// TIA Portal V19 export
// export: Created 2026-10-15T09:44:25.353626Z, ExportSetting WithDefaults, DisplayName Totally Integrated Automation Portal, DisplayVersion V19, DisplayName TIA Portal Openness, DisplayVersion V19, DisplayName TIA Portal Version Control Interface, DisplayVersion V19, DisplayName STEP 7 Professional, DisplayVersion V19, DisplayName STEP 7 Safety, DisplayVersion V19, DisplayName WinCC Basic/Comfort/Advanced, DisplayVersion V19, DisplayName WinCC Unified, DisplayVersion V19
FUNCTION "ROLL_WriteOutputs" : Void   // FC37, SCL
{ S7_Optimized_Access := 'TRUE' }
VERSION : 0.1
// stored: AutoNumber true, IsIECCheckEnabled false, SetENOAutomatically false, UDAEnableTagReadback false
   VAR_TEMP
      enabled : Bool;
   END_VAR
BEGIN

   IF "ROLL_IO".PhysicalIoConfigured THEN
       #enabled := "ROLL_IO".PhysicalOutputsEnabled AND NOT "ROLL_IO".Simulation AND NOT "ROLL_IO".ConversionFault;
       "Tag__639276542187652659" := #enabled AND "ROLL_IO".Output[16, 0];
       "Tag__639276542187732448" := #enabled AND "ROLL_IO".Output[16, 1];
       "Tag__639276542187792292" := #enabled AND "ROLL_IO".Output[16, 2];
       "Tag__639276542187852130" := #enabled AND "ROLL_IO".Output[16, 3];
       "Tag__639276542187911981" := #enabled AND "ROLL_IO".Output[16, 4];
       "Tag__639276542187972161" := #enabled AND "ROLL_IO".Output[16, 5];
       "Tag__639276542188021847" := #enabled AND "ROLL_IO".Output[16, 6];
       "Tag__639276542188081517" := #enabled AND "ROLL_IO".Output[16, 7];
       "Tag__639276542188141359" := #enabled AND "ROLL_IO".Output[17, 0];
       "Tag__639276542188191229" := #enabled AND "ROLL_IO".Output[17, 1];
       "Tag__639276542188251067" := #enabled AND "ROLL_IO".Output[17, 2];
       "Tag__639276542188320878" := #enabled AND "ROLL_IO".Output[17, 3];
       "Tag__639276542188410640" := #enabled AND "ROLL_IO".Output[17, 4];
       "Tag__639276542188520372" := #enabled AND "ROLL_IO".Output[17, 5];
       "Tag__639276542188610120" := #enabled AND "ROLL_IO".Output[17, 6];
       "Tag__639276542188699865" := #enabled AND "ROLL_IO".Output[17, 7];
       "Tag__639276542188769683" := #enabled AND "ROLL_IO".Output[18, 0];
       "Tag__639276542188839495" := #enabled AND "ROLL_IO".Output[18, 1];
       "Tag__639276542188899332" := #enabled AND "ROLL_IO".Output[18, 2];
       "Tag__639276542188969166" := #enabled AND "ROLL_IO".Output[18, 3];
       "Tag__639276542189049062" := #enabled AND "ROLL_IO".Output[18, 4];
       "Tag__639276542189108777" := #enabled AND "ROLL_IO".Output[18, 5];
       "Tag__639276542189178592" := #enabled AND "ROLL_IO".Output[18, 6];
       "Tag__639276542189258389" := #enabled AND "ROLL_IO".Output[18, 7];
       "Tag__639276542189338210" := #enabled AND "ROLL_IO".Output[19, 0];
       "Tag__639276542189407977" := #enabled AND "ROLL_IO".Output[19, 1];
       "Tag__639276542189488068" := #enabled AND "ROLL_IO".Output[19, 2];
       "Tag__639276542189557576" := #enabled AND "ROLL_IO".Output[19, 3];
       "Tag__639276542189627382" := #enabled AND "ROLL_IO".Output[19, 4];
       "Tag__639276542189697203" := #enabled AND "ROLL_IO".Output[19, 5];
       "Tag__639276542189767112" := #enabled AND "ROLL_IO".Output[19, 6];
       "Tag__639276542189836826" := #enabled AND "ROLL_IO".Output[19, 7];
       "Tag__639276542189916614" := #enabled AND "ROLL_IO".Output[20, 0];
       "Tag__639276542189996407" := #enabled AND "ROLL_IO".Output[20, 1];
       "Tag__639276542190076190" := #enabled AND "ROLL_IO".Output[20, 2];
       "Tag__639276542190146259" := #enabled AND "ROLL_IO".Output[20, 3];
       "Tag__639276542190215815" := #enabled AND "ROLL_IO".Output[20, 4];
       "Tag__639276542190295600" := #enabled AND "ROLL_IO".Output[20, 5];
       "Tag__639276542190365408" := #enabled AND "ROLL_IO".Output[20, 6];
       "Tag__639276542190435229" := #enabled AND "ROLL_IO".Output[20, 7];
       "Tag__639276542190505050" := #enabled AND "ROLL_IO".Output[21, 0];
       "Tag__639276542190574853" := #enabled AND "ROLL_IO".Output[21, 1];
       "Tag__639276542190654646" := #enabled AND "ROLL_IO".Output[21, 2];
       "Tag__639276542190724459" := #enabled AND "ROLL_IO".Output[21, 3];
       "Tag__639276542190804229" := #enabled AND "ROLL_IO".Output[21, 4];
       "Tag__639276542190874055" := #enabled AND "ROLL_IO".Output[21, 5];
       "Tag__639276542190943868" := #enabled AND "ROLL_IO".Output[21, 6];
       "Tag__639276542191023653" := #enabled AND "ROLL_IO".Output[21, 7];
       "Tag__639276542191093472" := #enabled AND "ROLL_IO".Output[22, 0];
       "Tag__639276542191173254" := #enabled AND "ROLL_IO".Output[22, 1];
       "Tag__639276542191253037" := #enabled AND "ROLL_IO".Output[22, 2];
       "Tag__639276542191332825" := #enabled AND "ROLL_IO".Output[22, 3];
       "Tag__639276542191402638" := #enabled AND "ROLL_IO".Output[22, 4];
       "Tag__639276542191482423" := #enabled AND "ROLL_IO".Output[22, 5];
       "Tag__639276542191552238" := #enabled AND "ROLL_IO".Output[22, 6];
       "Tag__639276542191612229" := #enabled AND "ROLL_IO".Output[22, 7];
       "Tag__639276542191672171" := #enabled AND "ROLL_IO".Output[23, 0];
       "Tag__639276542191731760" := #enabled AND "ROLL_IO".Output[23, 1];
       "Tag__639276542191791592" := #enabled AND "ROLL_IO".Output[23, 2];
       "Tag__639276542191841458" := #enabled AND "ROLL_IO".Output[23, 3];
       "Tag__639276542191901298" := #enabled AND "ROLL_IO".Output[23, 4];
       "Tag__639276542191951165" := #enabled AND "ROLL_IO".Output[23, 5];
       "Tag__639276542192011013" := #enabled AND "ROLL_IO".Output[23, 6];
       "Tag__639276542192070845" := #enabled AND "ROLL_IO".Output[23, 7];
       "Tag__639276542192120711" := #enabled AND "ROLL_IO".Output[24, 0];
       "Tag__639276542192180551" := #enabled AND "ROLL_IO".Output[24, 1];
       "Tag__639276542192240399" := #enabled AND "ROLL_IO".Output[24, 2];
       "Tag__639276542192290265" := #enabled AND "ROLL_IO".Output[24, 3];
       "Tag__639276542192350097" := #enabled AND "ROLL_IO".Output[24, 4];
       "Tag__639276542192399963" := #enabled AND "ROLL_IO".Output[24, 5];
       "Tag__639276542192459803" := #enabled AND "ROLL_IO".Output[24, 6];
       "Tag__639276542192509678" := #enabled AND "ROLL_IO".Output[24, 7];
       "Tag__639276542192569509" := #enabled AND "ROLL_IO".Output[25, 0];
       "Tag__639276542192619385" := #enabled AND "ROLL_IO".Output[25, 1];
       "Tag__639276542192679216" := #enabled AND "ROLL_IO".Output[25, 2];
       "Tag__639276542192729083" := #enabled AND "ROLL_IO".Output[25, 3];
       "Tag__639276542192778949" := #enabled AND "ROLL_IO".Output[25, 4];
       "Tag__639276542192839026" := #enabled AND "ROLL_IO".Output[25, 5];
       "Tag__639276542192888657" := #enabled AND "ROLL_IO".Output[25, 6];
       "Tag__639276542192938522" := #enabled AND "ROLL_IO".Output[25, 7];
   END_IF;
END_FUNCTION
